(* Schneider Machine Expert - Basic project native_literal_series_eight_il_only, file version 3.0.0.0 *)
(* ProjectInformations: Name=New project *)

HARDWARE
  Cpu 0: TM200CE40T
  EthernetConfiguration: NetworkName=M200, IpAllocationMode=FixedAddress, IpAddress=0.0.0.0, SubnetMask=0.0.0.0
  SerialLineConfiguration: Baud=Baud19200, Parity=ParityEven, DataBits=DataBits8, StopBits=StopBits1, PhysicalMedium=PhysicalMediumRs485, TransmissionMode=TransmissionModeModbusRtu, SlaveId=1, Addressing=SlaveAddressing
  MastTask: UsePeriodScanMode=false, PeriodScan=100
  FastTask: Period=255
  CpuBehavior: StartingMode=StartAsPreviousState, AutoSaveRamOnEeprom=true, WatchdogPeriod=250

SYMBOLS  (address, symbol, comment, settings)

POU New POU
  (* SectionNumber=0 *)

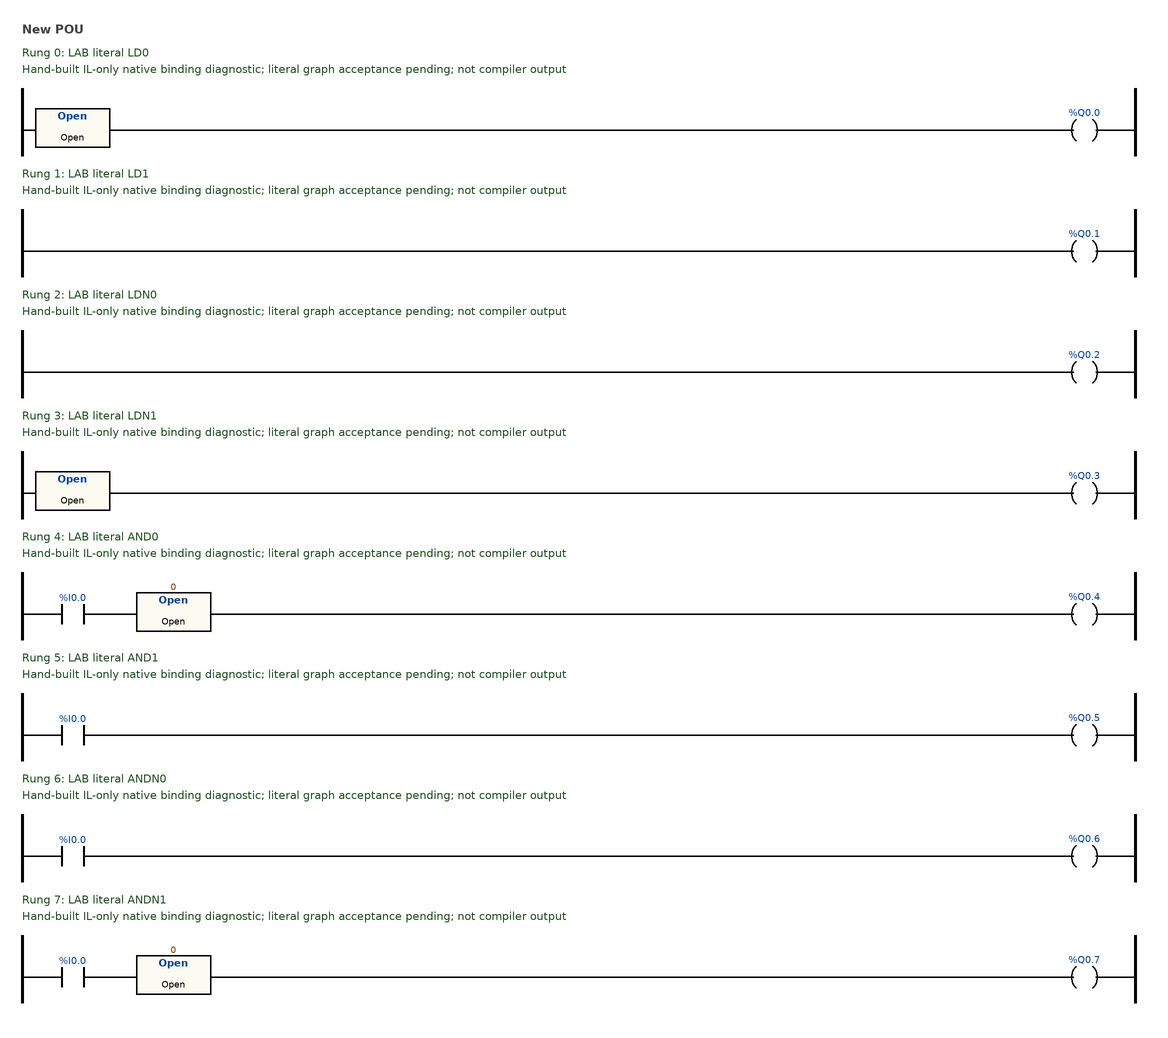

// Rung 0: LAB literal LD0
// Hand-built IL-only native binding diagnostic; literal graph acceptance pending; not compiler output
  LD 0
  ST %Q0.0
  // as ST:
  //   %Q0.0 := FALSE;

// Rung 1: LAB literal LD1
// Hand-built IL-only native binding diagnostic; literal graph acceptance pending; not compiler output
  LD 1
  ST %Q0.1
  // as ST:
  //   %Q0.1 := TRUE;

// Rung 2: LAB literal LDN0
// Hand-built IL-only native binding diagnostic; literal graph acceptance pending; not compiler output
  LD 1
  ST %Q0.2
  // as ST:
  //   %Q0.2 := TRUE;

// Rung 3: LAB literal LDN1
// Hand-built IL-only native binding diagnostic; literal graph acceptance pending; not compiler output
  LD 0
  ST %Q0.3
  // as ST:
  //   %Q0.3 := FALSE;

// Rung 4: LAB literal AND0
// Hand-built IL-only native binding diagnostic; literal graph acceptance pending; not compiler output
  LD %I0.0
  AND 0
  ST %Q0.4
  // as ST:
  //   %Q0.4 := %I0.0 AND FALSE;

// Rung 5: LAB literal AND1
// Hand-built IL-only native binding diagnostic; literal graph acceptance pending; not compiler output
  LD %I0.0
  AND 1
  ST %Q0.5
  // as ST:
  //   %Q0.5 := %I0.0;

// Rung 6: LAB literal ANDN0
// Hand-built IL-only native binding diagnostic; literal graph acceptance pending; not compiler output
  LD %I0.0
  AND 1
  ST %Q0.6
  // as ST:
  //   %Q0.6 := %I0.0;

// Rung 7: LAB literal ANDN1
// Hand-built IL-only native binding diagnostic; literal graph acceptance pending; not compiler output
  LD %I0.0
  AND 0
  ST %Q0.7
  // as ST:
  //   %Q0.7 := %I0.0 AND FALSE;
